(* IEC 61131-3 sources: codesys-to-astra/cds2astra/tests/corpus/C2A-LANG-OOP/neg/src/POUs/FB_A, 1 file *)

(* ---- FB_A.decl.st ---- *)
// Назначение: корпус правила cds2astra (synthetic).
// Автор:      kr0nsch
// Версия:     0.1.0
// Документ:   docs/RULES.md
FUNCTION_BLOCK FB_A
VAR
END_VAR
